FUNCTION_BLOCK AtvMedidasGen (* Medidas do ATV600 por Modbus generico (INT da planilha V4.6) para REAL na unidade de engenharia *)
  (* Standard: 61499-2 *)
  (* Version 0.1, 12/11/2026, Hidryco, Hidryco, Hidryco 12/11/2026: RFRD 8604 rpm (1 rpm), OTR 3205 torque (0,1 %), OPR 3211 potencia (1 %), UOP 3208 tensao do motor (1 V). *)
  PACKAGE SE.Nereda;
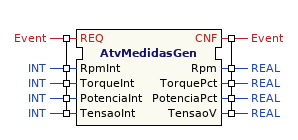
  EVENT_INPUT
    REQ WITH RpmInt, TorqueInt, PotenciaInt, TensaoInt; (* Converte *)
  END_EVENT
  EVENT_OUTPUT
    CNF WITH Rpm, TorquePct, PotenciaPct, TensaoV; (* Valores convertidos *)
  END_EVENT
  VAR_INPUT
    RpmInt : INT; (* RFRD 8604 - velocidade do motor (1 rpm) *)
    TorqueInt : INT; (* OTR 3205 - torque do motor (0,1 %) *)
    PotenciaInt : INT; (* OPR 3211 - potencia mecanica do motor (1 %) *)
    TensaoInt : INT; (* UOP 3208 - tensao do motor (1 V) *)
  END_VAR
  VAR_OUTPUT
    Rpm : REAL; (* Velocidade do motor (rpm) *)
    TorquePct : REAL; (* Torque do motor (%) *)
    PotenciaPct : REAL; (* Potencia do motor (%) *)
    TensaoV : REAL; (* Tensao do motor (V) *)
  END_VAR
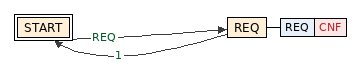
  EC_STATES
    START; (* Inicial *)
    REQ : REQ -> CNF; (* Converte *)
  END_STATES
  EC_TRANSITIONS
    START TO REQ := REQ;
    REQ TO START := 1;
  END_TRANSITIONS
  ALGORITHM REQ IN ST: (* Conversao *)
Rpm       := INT_TO_REAL(RpmInt);
TorquePct := INT_TO_REAL(TorqueInt) / 10.0;
PotenciaPct := INT_TO_REAL(PotenciaInt);
TensaoV   := INT_TO_REAL(TensaoInt);   (* UOP e UINT: ate 32767 V cabe em INT *)
  END_ALGORITHM
END_FUNCTION_BLOCK
